(* IEC 61131-3 sources: daoli-st-library/_quarantine, 3 files *)

(* ---- FC_DL_StatsRmsCalc.st ---- *)
(*==============================================================================
 * 组件名称 (Component)  : FC_DL_StatsRmsCalc
 * 所属子库 (Sublibrary) : DL_MathData
 * 当前版本 (Version)    : 1.0.0
 * 兼容性   (Platform)   : CODESYS 3.5+ / TwinCAT 3 / 汇川 InoProShop / 施耐德 Machine Expert
 *                         仅依赖 IEC 61131-3 标准数学（SQRT / ABS），零厂商私有库
 * 功能描述 (Function)   : 有效值 RMS 计算（交流量监测）：
 *                           RMS = SQRT( Σ x_i² / n )
 *                         与「均值」的本质差别：RMS 保留交流分量的能量（直流表读 0，
 *                         RMS 表读出真实有效值），故适用于电流/电压有效值、
 *                         振动加速度有效值、阀线圈 PWM 电流有效值的单批核算。
 *                         **溢出前置防护**：LREAL 可表到 1.8E308，故 |x| > 1E150 时
 *                         x² 会越过可表上限。本件在累加前先扫一遍最大绝对值，
 *                         超阈即判故障级 eOverflowRisk 并拒绝计算（不输出 Inf）。
 * 接口     (Interface)  : 输入 afSample 样本数组 [EU]、iCount 有效样本数 [个]（1..64）；
 *                         输出 fRms 有效值 [EU]、fPeak 最大绝对值（峰值） [EU]、
 *                         fSumSq 平方和（诊断用） [EU^2]、bValid 结果可信、
 *                         eErrCode（E_DL_StatsRmsErr）；
 *                         返回值 = bValid。
 * 边界     (Boundary)   : ① 属主边界：只算单批 RMS，不做跨周期累计（跨周期归 FB）、
 *                         不做真有效值（含谐波分量的时域积分，需更高采样率）。
 *                         ② 样本数域闸 1..64；越域 → 故障级 eBadCount。
 *                         n=1 时 RMS = |x1|，合法。
 *                         ③ 非有限双判：全部有效样本逐项枚举。
 *                         ④ 溢出前置防护阈值 DL_SRC_MAG_MAX = 1E150（平方后 1E300，仍在 LREAL 域内）。
 *                         ⑤ 平方和与 RMS 均做非有限复检；RMS 必须 >= 0（负值判内部不一致）。
 *                         ⑥ 零全局耦合（无 GVL / VAR_EXTERNAL / 物理地址）。
 * 分工声明 (Scope)      : 与 `FC_DL_StatsMeanStdDev` 分工：均值/标准差（去直流）归那件、
 *                         含直流的有效值归本件；与 `FC_DL_StatsZeroCrossRate` 分工：
 *                         频率特征归那件。
 * 来源标签 (Source Tag) : 原创实现（无外部代码引入）
 * 码表     (Codes)      : 本件不占用全局数字码位；出口为 BOOL + 3×LREAL +
 *                         本文件内定义 enum E_DL_StatsRmsErr（全库唯一）。
 * 红线自检 (Redline)    : R1 ✓ 零 GVL/VAR_EXTERNAL ｜ R2 ✓ 零 %I/%Q/%M ｜ R3 ✓ 纯 IEC 61131-3
 *                         R4 ✓ 点数域闸 + 全样本非有限双判 + 平方溢出前置防护 + 结果复检 ｜ R5 ✓ 声明逐行同行双语注释
 *                         R6 N/A（纯函数无状态机） ｜ R7 N/A（无实例调用）
 * 修订历史 (Revision)   : 2026-11-23  v1.0.0  R77 首版（批次 B3 · 序号 19）
 * 验收向量 (Acceptance) : ① afSample=[3,4], iCount=2 → 平方和 25，RMS=SQRT(12.5)≈3.535533906
 *                         （容差 1E-9），fPeak=4.0；
 *                         ② afSample=[1,-1,1,-1], iCount=4 → 平方和 4，RMS=1.0（直流为 0 但 RMS 非 0）；
 *                         ③ afSample=[0,0,0], iCount=3 → fRms=0.0, fPeak=0.0, eOk；
 *                         ④ afSample=[1E200], iCount=1 → 返回 FALSE, eOverflowRisk（不输出 Inf）；
 *                         ⑤ iCount=65 → 返回 FALSE, eBadCount。
 *==============================================================================*)

(*-----------------------------------------------------------------------------
 * 枚举: E_DL_StatsRmsErr（有效值统计错误码，归属 DL_MathData，与本件同文件，全库唯一属主）
 *----------------------------------------------------------------------------*)
TYPE E_DL_StatsRmsErr :
(
    eOk           := 0,   // 信息级：计算完成 / Info: computed
    eBadCount     := 1,   // 故障级：样本数越域 / Fault: sample count out of domain
    eNonFinite    := 2,   // 故障级：样本含非有限值 / Fault: non-finite sample present
    eOverflowRisk := 3,   // 故障级：量值平方将越出可表域 / Fault: squaring would overflow the representable range
    eInternal     := 9    // 故障级：RMS 为负等内部不一致 / Fault: negative RMS or other internal inconsistency
);
END_TYPE

FUNCTION FC_DL_StatsRmsCalc : BOOL
VAR_INPUT
    afSample : ARRAY[1..64] OF LREAL;  // 样本数组 [EU] / Sample array
    iCount   : INT;                    // 有效样本数（1..64） [个] / Valid sample count, 1..64
END_VAR
VAR_OUTPUT
    fRms      : LREAL;  // 有效值 [EU] / Root mean square
    fPeak     : LREAL;  // 最大绝对值 [EU] / Peak absolute value
    fSumSq    : LREAL;  // 平方和（诊断用） [EU^2] / Sum of squares for diagnostics
    bValid    : BOOL;   // 结果可信标志 [-] / Result trustworthy flag
    eErrCode  : E_DL_StatsRmsErr; // 错误码出口 [-] / Error code outlet
END_VAR
VAR
    _i        : INT;    // 样本遍历下标 [-] / Sample index
    _bNonFin  : BOOL;   // 非有限标志 [-] / Non-finite flag
    _fAbs     : LREAL;  // 当前样本绝对值 [EU] / Current absolute value
    _fPeak    : LREAL;  // 最大绝对值累计 [EU] / Peak accumulator
    _fSumSq   : LREAL;  // 平方和累计 [EU^2] / Sum of squares accumulator
    _fMeanSq  : LREAL;  // 均方值 [EU^2] / Mean square value
END_VAR
VAR CONSTANT
    DL_SRC_CNT_MIN : INT := 1;          // 样本数下限 [个] / Count lower bound
    DL_SRC_CNT_MAX : INT := 64;         // 样本数上限（数组容量） [个] / Count upper bound
    DL_SRC_MAG_MAX : LREAL := 1.0E150;  // 平方溢出前置阈值（平方后 1E300 仍可表） [EU] / Pre-square overflow threshold
    DL_SRC_ZERO    : LREAL := 0.0;      // 零基准（含非有限判零） [-] / Zero base including non-finite probe
END_VAR

(* —— 段 0：出口预置安全值 —— *)
FC_DL_StatsRmsCalc := FALSE;                       // 返回值预置无效 / Return preset invalid
fRms     := DL_SRC_ZERO;                           // RMS 哨兵 / RMS sentinel
fPeak    := DL_SRC_ZERO;                           // 峰值哨兵 / Peak sentinel
fSumSq   := DL_SRC_ZERO;                           // 平方和哨兵 / Sum of squares sentinel
bValid   := FALSE;                                 // 可信标志预置否 / Trust flag preset false
eErrCode := E_DL_StatsRmsErr.eBadCount;            // 预置最严码 / Preset strictest code

(* —— 段 1：样本数域闸 —— *)
IF (iCount < DL_SRC_CNT_MIN) OR (iCount > DL_SRC_CNT_MAX) THEN
    RETURN;
END_IF

(* —— 段 2：非有限域闸 + 量值上限扫描（平方溢出前置防护，一遍完成两件事） —— *)
_bNonFin := FALSE;
_fPeak   := DL_SRC_ZERO;
_i := 1;
WHILE _i <= iCount DO
    IF (afSample[_i] <> afSample[_i]) OR ((afSample[_i] - afSample[_i]) <> DL_SRC_ZERO) THEN
        _bNonFin := TRUE;                          // 样本非有限 / Sample non-finite
    ELSE
        _fAbs := ABS(afSample[_i]);                // 绝对值 / Absolute value
        IF _fAbs > _fPeak THEN
            _fPeak := _fAbs;                       // 更新峰值 / Update peak
        END_IF
    END_IF
    _i := _i + 1;
END_WHILE
IF _bNonFin THEN
    eErrCode := E_DL_StatsRmsErr.eNonFinite;       // 故障级码 / Fault-level code
    RETURN;
END_IF
IF _fPeak > DL_SRC_MAG_MAX THEN
    eErrCode := E_DL_StatsRmsErr.eOverflowRisk;    // 故障级：平方将溢出 / Fault: squaring would overflow
    RETURN;                                        // 拒绝计算，绝不输出 Inf / Refuse rather than emit Inf
END_IF

(* —— 段 3：平方和累加 —— *)
_fSumSq := DL_SRC_ZERO;
_i := 1;
WHILE _i <= iCount DO
    _fSumSq := _fSumSq + afSample[_i] * afSample[_i];   // 逐点平方累加 / Accumulate squares
    _i := _i + 1;
END_WHILE

(* —— 段 4：均方与 RMS（分母 n 已由段 1 保证 >= 1，无除零） —— *)
_fMeanSq := _fSumSq / INT_TO_LREAL(iCount);        // 均方值 / Mean square
fRms     := SQRT(_fMeanSq);                        // 有效值 / Root mean square

(* —— 段 5：结果复检（非有限 + 非负 + 不超峰值） —— *)
IF (fRms <> fRms) OR (_fSumSq <> _fSumSq) THEN
    fRms     := DL_SRC_ZERO;                       // 复检异常回哨兵 / Recheck failed: sentinel
    fSumSq   := DL_SRC_ZERO;
    fPeak    := DL_SRC_ZERO;
    eErrCode := E_DL_StatsRmsErr.eNonFinite;
    RETURN;
END_IF
IF (fRms < DL_SRC_ZERO) OR (fRms > _fPeak) THEN
    fRms     := DL_SRC_ZERO;                       // RMS 必在 [0, peak] 内，否则内部不一致 / RMS must lie in 0..peak
    fSumSq   := DL_SRC_ZERO;
    fPeak    := DL_SRC_ZERO;
    eErrCode := E_DL_StatsRmsErr.eInternal;
    RETURN;
END_IF

(* —— 段 6：成功出口 —— *)
fSumSq   := _fSumSq;                               // 导出平方和 / Export sum of squares
fPeak    := _fPeak;                                // 导出峰值 / Export peak
bValid   := TRUE;
eErrCode := E_DL_StatsRmsErr.eOk;                  // 信息级成功 / Info success
FC_DL_StatsRmsCalc := TRUE;                        // 结果可信 / Result trustworthy

END_FUNCTION

(* ---- FC_DL_StringPadLeftZeros.st ---- *)
(*==============================================================================
 * 组件名称 (Component)  : FC_DL_StringPadLeftZeros
 * 所属子库 (Sublibrary) : DL_Base
 * 当前版本 (Version)    : 1.0.0
 * 兼容性   (Platform)   : CODESYS 3.5+ / TwinCAT 3 / 汇川 InoProShop / 施耐德 Machine Expert
 *                         仅依赖 IEC 61131-3 标准字符串九函数（LEN / LEFT / CONCAT），零厂商私有库
 * 功能描述 (Function)   : 左补零至定长（编号 / 时间戳 / 批号规范化）。
 *                         sIn 左侧填充 pad 字符（默认 '0'）至 uiTargetLen 长度；
 *                         sIn 已达或超过目标长度时原样返回（不截断）并置 bOverflow；
 *                         目标长度超过缓冲上限 255 时钳位至 255 并置 bOverflow。
 *                         用于 PLC 侧生成定宽字符串键（如 "00042"），便于 HMI 对齐与
 *                         上位机字典排序（定宽字典序 = 数值序）。
 * 接口     (Interface)  : 输入 sIn 原始字符串 [-]、uiTargetLen 目标定长 [字符]、
 *                         sPadChar 填充字符（取首字符，空串视为 '0'）[-]；
 *                         输出 sOut 结果字符串、uiOutLen 实际字符数 [字符]、
 *                         bOverflow 溢出/钳位回执、eErrCode 错误码（E_DL_StrPadErr）；
 *                         返回值 = bValid 转换有效标志（TRUE = sOut 可信）。
 * 边界     (Boundary)   : ① 属主边界：只做补位，不做数值格式化、不做千分位、不截断。
 *                         ② 全局缓冲上限 255（STRING(255) 契约），目标超限钳位并置
 *                         bOverflow（信息级码 eClampLen，不置故障）。
 *                         ③ 输入为空串时输出全填充串（长度 = uiTargetLen），合法。
 *                         ④ 索引全 1 基（IEC 字符串函数约定），无 0 基偏移路径。
 *                         ⑤ 零全局耦合（无 GVL / VAR_EXTERNAL / 物理地址）。
 * 分工声明 (Scope)      : 与 `FC_DL_StringTruncEllipsis` 分工：超长截断归那件，
 *                         本件超长只回执不截断（补位与截断语义互斥，避免隐式改写）。
 *                         与 `FC_DL_StringRepeat` 分工：重复拼接归那件，本件只补单字符。
 * 来源标签 (Source Tag) : 原创实现（无外部代码引入）
 * 码表     (Codes)      : 本件不占用全局数字码位；出口为 BOOL 返回 + STRING 结果 +
 *                         本文件内定义 enum E_DL_StrPadErr（全库唯一）。
 * 红线自检 (Redline)    : R1 ✓ 零 GVL/VAR_EXTERNAL ｜ R2 ✓ 零 %I/%Q/%M ｜ R3 ✓ 纯 IEC 61131-3
 *                         R4 ✓ 目标长度双侧钳位 + 循环上限硬保护 ｜ R5 ✓ 声明逐行同行双语注释
 *                         R6 N/A（纯函数无状态机） ｜ R7 N/A（无实例调用）
 * 修订历史 (Revision)   : 2026-11-23  v1.0.0  R77 首版（批次 B2 · 序号 1）
 * 验收向量 (Acceptance) : ① sIn='42', uiTargetLen=5, sPadChar='0' → sOut='00042',
 *                         uiOutLen=5, bOverflow=FALSE, 返回 TRUE, eErrCode=eOk；
 *                         ② sIn='123456', uiTargetLen=3 → sOut='123456'（原样不截断）,
 *                         uiOutLen=6, bOverflow=TRUE, 返回 TRUE, eErrCode=eOverflowInput；
 *                         ③ sIn='', uiTargetLen=3 → sOut='000', uiOutLen=3, eOk；
 *                         ④ uiTargetLen=300 → 钳位 255，bOverflow=TRUE, eClampLen。
 *==============================================================================*)

(*-----------------------------------------------------------------------------
 * 枚举: E_DL_StrPadErr（左补零错误码，归属 DL_Base，与本件同文件，全库唯一属主）
 * 分级: 故障级码（eInvalidParam）恒伴返回 FALSE；信息级码（eOk / eOverflowInput /
 *       eClampLen）返回 TRUE 且结果仍可信。
 *----------------------------------------------------------------------------*)
TYPE E_DL_StrPadErr :
(
    eOk            := 0,   // 信息级：正常补位完成 / Info: padding completed
    eOverflowInput := 1,   // 信息级：输入已达目标长度，原样返回 / Info: input already long enough, returned as-is
    eClampLen      := 2,   // 信息级：目标长度超缓冲上限已钳位 / Info: target length clamped to buffer ceiling
    eInvalidParam  := 3    // 故障级：参数非法（填充串全空且目标长度非正） / Fault: invalid parameter
);
END_TYPE

FUNCTION FC_DL_StringPadLeftZeros : BOOL
VAR_INPUT
    sIn         : STRING(255);   // 原始字符串（待补位） [-] / Raw input string to be padded
    uiTargetLen : UINT;          // 目标定长，合法域 1..255 [字符] / Target fixed length, domain 1..255 [chars]
    sPadChar    : STRING(255);   // 填充字符源（取首字符，空串按 '0'） [-] / Pad character source, first char, empty means '0'
END_VAR
VAR_OUTPUT
    sOut        : STRING(255);   // 补位结果字符串 [-] / Padded result string
    uiOutLen    : UINT;          // 结果实际字符数 [字符] / Actual character count of result [chars]
    bOverflow   : BOOL;          // 溢出/钳位回执（信息级，不置故障） [-] / Overflow or clamp receipt, info level
    eErrCode    : E_DL_StrPadErr; // 错误码出口 [-] / Error code outlet
END_VAR
VAR
    _uiInLen    : UINT;          // 输入字符串字符数 [字符] / Input character count [chars]
    _uiPadNum   : UINT;          // 需补入的填充字符个数 [字符] / Number of pad characters required [chars]
    _sPadOne    : STRING(255);   // 单字符填充串（循环拼接基元） [-] / Single-character pad unit for concatenation
    _i          : UINT;          // 填充循环计数器 [-] / Padding loop counter
END_VAR
VAR CONSTANT
    DL_SPZ_LEN_MAX : UINT := 255;   // 缓冲上限（STRING(255) 契约） [字符] / Buffer ceiling per STRING(255) contract [chars]
    DL_SPZ_LEN_MIN : UINT := 1;     // 目标长度下限（0 视为非法参数） [字符] / Target length lower bound, 0 is invalid [chars]
    DL_SPZ_ZERO_CH : STRING(255) := '0'; // 默认填充字符 / Default pad character
END_VAR

(* —— 段 0：出口预置安全值（预置最严码 + 哨兵输出） —— *)
FC_DL_StringPadLeftZeros := FALSE;                // 返回值预置无效 / Return preset invalid
sOut      := '';                                  // 结果哨兵空串 / Result sentinel empty string
uiOutLen  := 0;                                   // 长度哨兵 0 / Length sentinel zero
bOverflow := FALSE;                               // 溢出口预置正常 / Overflow preset normal
eErrCode  := E_DL_StrPadErr.eInvalidParam;        // 预置最严码，参数闸命中直接早退 / Preset strictest code

(* —— 段 1：参数域闸（目标长度下限；分母型参数无，纯域判定） —— *)
IF uiTargetLen < DL_SPZ_LEN_MIN THEN
    RETURN;                                       // 目标长度 0：保持故障码与哨兵 / Zero target length: keep fault code
END_IF

(* —— 段 2：目标长度上限钳位（缓冲可表性反算，R 饱和硬限） —— *)
IF uiTargetLen > DL_SPZ_LEN_MAX THEN
    uiTargetLen := DL_SPZ_LEN_MAX;                 // 钳位至缓冲上限 / Clamp to buffer ceiling
    bOverflow   := TRUE;                           // 钳位回执 / Clamp receipt
    eErrCode    := E_DL_StrPadErr.eClampLen;       // 信息级码 / Info-level code
END_IF

(* —— 段 3：输入长度实测（LEN 返回 UDINT，标准函数显式收窄到 UINT） —— *)
_uiInLen := UDINT_TO_UINT(LEN(sIn));               // 输入字符数 / Input character count

(* —— 段 4：已达目标长度：原样返回不截断（早退分支，语义显式） —— *)
IF _uiInLen >= uiTargetLen THEN
    sOut      := sIn;                              // 原样返回 / Return as-is
    uiOutLen  := _uiInLen;                         // 实际长度取输入长度 / Length equals input length
    bOverflow := TRUE;                             // 已达/超过目标长度回执 / Already at or beyond target
    eErrCode  := E_DL_StrPadErr.eOverflowInput;    // 信息级码（覆盖钳位码，更贴语义） / Info code overrides clamp code
    FC_DL_StringPadLeftZeros := TRUE;              // 结果可信 / Result trustworthy
    RETURN;                                        // 早退 / Early exit
END_IF

(* —— 段 5：填充字符解析（空串按默认 '0'，否则取首字符） —— *)
IF LEN(sPadChar) = 0 THEN
    _sPadOne := DL_SPZ_ZERO_CH;                    // 空串回落默认字符 / Empty falls back to default character
ELSE
    _sPadOne := LEFT(sPadChar, 1);                 // 取首字符（1 基索引） / Take first character, 1-based
END_IF

(* —— 段 6：循环左补（补数已由上限钳位保证 <= 255，循环有界） —— *)
_uiPadNum := uiTargetLen - _uiInLen;               // 需补个数 = 目标 - 现有 / Pad count = target - existing
sOut      := _sPadOne;                             // 以单个填充字符起头，避免首次拼接空串副作用 / Start with one pad unit
IF _uiPadNum > DL_SPZ_LEN_MIN THEN
    FOR _i := 2 TO _uiPadNum DO
        sOut := CONCAT(sOut, _sPadOne);            // 逐个追加填充字符 / Append one pad character per iteration
    END_FOR;
END_IF
sOut := CONCAT(sOut, sIn);                         // 左补齐后接原串 / Append original string after pad prefix

(* —— 段 7：结果复检（长度必须等于目标，否则判内部不一致） —— *)
uiOutLen := UDINT_TO_UINT(LEN(sOut));              // 实测结果长度 / Measured result length
IF uiOutLen <> uiTargetLen THEN
    sOut     := '';                                // 复检失败回哨兵 / Recheck failed: back to sentinel
    uiOutLen := 0;                                 // 长度回哨兵 / Length back to sentinel
    eErrCode := E_DL_StrPadErr.eInvalidParam;      // 故障级码 / Fault-level code
    RETURN;                                        // 返回 FALSE 保持 / Keep return FALSE
END_IF

(* —— 段 8：成功出口（信息级码保留，bOverflow 供调用方判别） —— *)
IF eErrCode = E_DL_StrPadErr.eClampLen THEN
    bOverflow := TRUE;                             // 钳位情形回执保持 / Keep clamp receipt
END_IF
FC_DL_StringPadLeftZeros := TRUE;                  // 补位有效 / Padding valid

END_FUNCTION

(* ---- FB_DL_RunningAverageN.st ---- *)
(*==============================================================================
 * 组件名称 (Component)  : FB_DL_RunningAverageN
 * 所属子库 (Sublibrary) : DL_Algo
 * 当前版本 (Version)    : 1.0.0
 * 兼容性   (Platform)   : CODESYS 3.5+ / TwinCAT 3 / 汇川 InoProShop / 施耐德 Machine Expert
 *                         仅依赖 IEC 61131-3（INT_TO_LREAL），零厂商私有库
 * 功能描述 (Function)   : N 点滑动均值（环形缓冲，增量求和）。窗口 N 可配 1..32，
 *                         运行中变更窗口自动清表重建（避免新旧两段样本混算）。
 *                         算法：写入前先减去被覆盖的最老样本（_fSum := _fSum - old + new），
 *                         均值 = _fSum / 当前样本数，故单拍开销与 N 无关（O(1)）。
 *                         用途：编码器速度、流量、称重等周期性抖动量平滑。
 * 接口     (Interface)  : 输入 bEnable 使能、bReset 清表复位、fIn 采样输入 [EU]、
 *                         iWindow 窗口点数 [个]（1..32）；
 *                         输出 fOut 均值 [EU]、iFillCount 当前样本数 [个]、
 *                         bValid 输出有效、bError 故障标志、uErrorId 故障码；
 *                         返回值由 FB 实例状态提供（无返回值，读 bValid）。
 * 边界     (Boundary)   : ① 属主边界：只做算术均值，不做中值 / 加权 / 剔除离群（另件）。
 *                         ② 非有限输入 → 进故障态、**冻结输出**（不更新），uErrorId=16#0003_0002；
 *                         故障态只能由 bEnable=FALSE 或 bReset 解除（可达恢复路径）。
 *                         ③ 窗口域闸 1..32：越域钳位并置信息码 16#0003_0001，不中断扫描。
 *                         ④ 除零防护：均值除法前判 _iFill >= 1。
 *                         ⑤ 零全局耦合（无 GVL / VAR_EXTERNAL / 物理地址）。
 * 分工声明 (Scope)      : 与 `FB_DL_LowPassFilter` 分工：一阶惯性归那件（无限记忆）、
 *                         有限窗口算术均值归本件；与统计族 FC 分工：一次性批统计归 FC。
 * 来源标签 (Source Tag) : 原创实现（无外部代码引入）
 * 码表     (Codes)      : 16#0003_0000 无故障 / 16#0003_0001 窗口越域已钳位（信息级）/
 *                         16#0003_0002 输入非有限（故障级）/ 16#0003_0005 非法状态（故障级）。
 * 红线自检 (Redline)    : R1 ✓ 零 GVL/VAR_EXTERNAL ｜ R2 ✓ 零 %I/%Q/%M ｜ R3 ✓ 纯 IEC 61131-3
 *                         R4 ✓ 除零前置判零 + 窗口域闸 + 非有限拒绝 ｜ R5 ✓ 声明逐行同行双语注释
 *                         R6 ✓ 四态 ENUM + CASE + ELSE 兜底 ｜ R7 N/A（无 TON/边沿实例）
 * 修订历史 (Revision)   : 2026-11-23  v1.0.0  R77 首版（批次 B3 · 序号 9）
 * 验收向量 (Acceptance) : ① iWindow=4，依次输入 1,2,3,4,5 → 第 4 拍 fOut=2.5；
 *                         第 5 拍（窗口已满，挤掉 1）→ fOut=(2+3+4+5)/4=3.5；
 *                         ② bReset=TRUE 一拍 → iFillCount=0，fOut=0.0，bValid=FALSE；
 *                         ③ iWindow=0 → 钳位为 1，uErrorId=16#0003_0001，仍正常输出；
 *                         ④ fIn=NaN → uErrorId=16#0003_0002，bError=TRUE，fOut 冻结上拍值；
 *                         ⑤ iWindow=40 → 钳位 32，uErrorId=16#0003_0001。
 *==============================================================================*)

(*-----------------------------------------------------------------------------
 * 枚举: E_DL_RavgState（滑动均值状态机，归属 DL_Algo，与本件同文件，全库唯一属主）
 *----------------------------------------------------------------------------*)
TYPE E_DL_RavgState :
(
    eInit  := 0,    // 首扫 / 复位后：清表并直取首个样本 / First scan or after reset: clear and seed
    eRun   := 10,   // 运行态：环形缓冲增量均值 / Running: incremental ring-buffer average
    eHold   := 20,  // 保持态：未使能，输出冻结 / Hold: disabled, output frozen
    eFault := 99    // 故障态：输出冻结，等待 bEnable 跌落或 bReset / Fault: frozen, awaiting disable or reset
);
END_TYPE

FUNCTION_BLOCK FB_DL_RunningAverageN
VAR_INPUT
    bEnable : BOOL := FALSE;   // 使能，FALSE 冻结输出 / Enable, FALSE freezes output
    bReset  : BOOL := FALSE;   // 复位清表（单拍有效） / Reset and clear buffer, single scan
    fIn     : LREAL := 0.0;    // 采样输入 [EU] / Sampling input [EU]
    iWindow : INT := 8;        // 窗口点数，合法域 1..32 [个] / Window size, domain 1..32
END_VAR
VAR_OUTPUT
    fOut       : LREAL;   // 滑动均值输出 [EU] / Moving average output [EU]
    iFillCount : INT;     // 当前有效样本数 [个] / Current valid sample count
    bValid     : BOOL;    // 输出有效标志 [-] / Output valid flag
    bError     : BOOL;    // 故障标志，与 uErrorId 联动 [-] / Fault flag coupled with uErrorId
    uErrorId   : UDINT;   // 故障码，0 = 无故障 [-] / Error code, zero means healthy
END_VAR
VAR
    _afBuf   : ARRAY[1..32] OF LREAL;  // 环形样本缓冲 [EU] / Ring sample buffer
    _fSum    : LREAL;                  // 样本和（增量维护） [EU] / Sample sum maintained incrementally
    _iHead   : INT;                    // 环形写入位（最老样本位） [-] / Ring write position, oldest slot
    _iFill   : INT;                    // 当前样本数 [个] / Current sample count
    _iWinEff : INT;                    // 生效窗口（钳位后） [个] / Effective window after clamping
    _i       : INT;                    // 循环下标 [-] / Loop index
    eState   : E_DL_RavgState;         // 状态机当前状态 [-] / Current state
END_VAR
VAR CONSTANT
    DL_RAV_WIN_MIN : INT := 1;       // 窗口下限 [个] / Window lower bound
    DL_RAV_WIN_MAX : INT := 32;      // 窗口上限（数组容量） [个] / Window upper bound
    DL_RAV_ZERO_L  : LREAL := 0.0;   // 零基准（含非有限判零） [-] / Zero base including non-finite probe
END_VAR

(* —— 段 1：参数域闸（不中断扫描，只钳位并置信息码） —— *)
uErrorId := 16#0003_0000;                          // 预置无故障 / Preset healthy
_iWinEff := iWindow;
IF iWindow < DL_RAV_WIN_MIN THEN
    _iWinEff := DL_RAV_WIN_MIN;                    // 窗口过小钳位 / Too small window clamped
    uErrorId := 16#0003_0001;                      // 信息级：窗口越域已钳位 / Info: window clamped
ELSIF iWindow > DL_RAV_WIN_MAX THEN
    _iWinEff := DL_RAV_WIN_MAX;                    // 窗口过大钳位 / Too large window clamped
    uErrorId := 16#0003_0001;                      // 信息级：窗口越域已钳位 / Info: window clamped
END_IF

(* —— 段 2：非有限输入防御（进故障态冻结输出，最短恢复路径 = bEnable 跌落或 bReset） —— *)
IF (fIn <> fIn) OR ((fIn - fIn) <> DL_RAV_ZERO_L) THEN
    eState   := eFault;                            // 强制故障态 / Force fault state
    uErrorId := 16#0003_0002;                      // 故障级：输入非有限 / Fault: non-finite input
END_IF

(* —— 段 3：窗口变更或复位 → 回首扫态（清表重建） —— *)
IF bReset THEN
    eState := eInit;                               // 复位请求回首扫 / Reset request returns to init
END_IF

(* —— 段 4：状态派生（故障态保持；未使能保持；其余运行） —— *)
IF NOT bEnable THEN
    eState := eHold;                               // 未使能：保持并冻结输出 / Disabled: hold and freeze
ELSIF eState = eFault THEN
    eState := eFault;                              // 故障态保持，等待外部解除 / Fault holds until cleared
ELSIF eState = eInit THEN
    eState := eInit;                               // 首扫态保持一拍 / Init holds for one scan
ELSE
    eState := eRun;                                // 常规运行 / Normal running
END_IF

(* —— 段 5：主状态机（CASE 覆盖 + ELSE 兜底） —— *)
CASE eState OF

    eInit:
        (* 清表：缓冲、求和、指针、计数全部归零，再以本拍样本播种（避免首拍均值 = 0） *)
        FOR _i := 1 TO DL_RAV_WIN_MAX DO
            _afBuf[_i] := DL_RAV_ZERO_L;
        END_FOR;
        _fSum    := DL_RAV_ZERO_L;
        _iFill   := 1;                             // 播种首个样本 / Seed first sample
        _iHead   := 1;
        _afBuf[1] := fIn;
        _fSum    := fIn;
        fOut     := fIn;                           // 首拍直取样本，无历史瞬态 / First scan follows input
        bValid   := TRUE;
        eState   := eRun;                          // 下一拍进入运行态 / Move to running next scan

    eRun:
        IF _iFill < _iWinEff THEN
            (* 未满窗：追加写入（无样本被挤出） *)
            _iFill := _iFill + 1;
            _iHead := _iFill;
            _afBuf[_iHead] := fIn;
            _fSum  := _fSum + fIn;
        ELSE
            (* 满窗：先减去被覆盖的最老样本，再写入新样本（增量 O(1)） *)
            _fSum := _fSum - _afBuf[_iHead] + fIn;
            _afBuf[_iHead] := fIn;
            _iHead := _iHead + 1;                  // 写入位前移 / Advance write slot
            IF _iHead > _iWinEff THEN
                _iHead := 1;                       // 环形回绕 / Wrap around
            END_IF
        END_IF
        IF _iFill >= 1 THEN
            fOut := _fSum / INT_TO_LREAL(_iFill);  // 除零已判（_iFill >= 1） / Division guarded
        ELSE
            fOut := DL_RAV_ZERO_L;                 // 防御兜底（结构上不可达） / Defensive fallback
        END_IF
        bValid := TRUE;

    eHold:
        (* 未使能：输出冻结保持上拍值，样本表不变，恢复使能后继续累积 *)
        (* Disabled: output frozen, buffer untouched, accumulation resumes on enable *)
        bValid := FALSE;

    eFault:
        (* 故障态：输出冻结保持上拍值（不推到 0，避免下游误判为真实零值） *)
        (* Fault: output frozen rather than zeroed, so downstream sees no fake zero *)
        bValid := FALSE;

    ELSE
        (* 非法状态拦截：任何未定义枚举值一律进故障态并置公共兜底码 *)
        eState   := eFault;
        bValid   := FALSE;
        uErrorId := 16#0003_0005;                  // 故障级：非法状态 / Fault: illegal state

END_CASE;

(* —— 段 6：出口映射（名实双出口：bError 与 uErrorId 同源） —— *)
iFillCount := _iFill;                              // 导出当前样本数 / Export sample count
bError     := (uErrorId <> 16#0003_0000);          // 故障级码才置 bError（信息级 16#0003_0001 不置） / Fault-level only

END_FUNCTION_BLOCK
